(*
SPDX-FileCopyrightText: © 2026 Oleksandr Tiutyk <trofimich@gmail.com>
SPDX-License-Identifier: MIT
License: https://opensource.org/license/mit
*)

(*! <summary>Orders the top-level runner calls and publication of their observations.</summary> *)
{attribute 'qualified_only'}
{attribute 'strict'}
TYPE RUNNER_TEST_PHASE :
(
	CHECK_CONSTRUCTION,
	INITIALIZE_ROOTS,
	EXECUTE_ROOTS,
	CHECK_NULL_ROOT,
	CHECK_EMPTY_ROOTS,
	CHECK_DUPLICATE_ROOT,
	PUBLISH_RESULTS,
	FINISHED
);
END_TYPE

(* stored: Version 1.1.0.1
   DUT RUNNER_TEST_PHASE: Id {0fc9fc44-302e-4d89-a860-003934491678} *)
